Fanuc KAREL source: KX00018.KL

PROGRAM KX00018
%NOLOCKGROUP
VAR
  I: INTEGER
  J: INTEGER
  B: BOOLEAN
  F: FILE
  S: STRING[80]
  P: XYZWPR
  BA: ARRAY[4] OF BYTE
BEGIN
  BA[1] = 7
  I = BA[1]
END KX00018
